Fanuc KAREL source: KC00028.KL

PROGRAM KC00028
%NOLOCKGROUP
%ENVIRONMENT MOTN
VAR
  I: INTEGER
  J: INTEGER
  K: INTEGER
  R: REAL
  B: BOOLEAN
  S: STRING[80]
  T: STRING[80]
  P: PATH
  Q: PATH
  AI: ARRAY[8] OF INTEGER
  AB: ARRAY[244] OF BYTE
  JP: JOINTPOS
  P1: POSITION
  P2: POSITION
  P3: POSITION
  C: CONFIG
  AR: ARRAY[9] OF REAL
BEGIN
  POS2JOINT(JP,P1,P2,P3,I,C,AR,JP,J)
END KC00028
